// TIA Portal V20 export
DATA_BLOCK "POS3_0_Signal"   // DB34
{ S7_Optimized_Access := 'TRUE' }
// stored: MemoryReserve 100
   VAR
      Schrittkette { S7_SetPoint := 'True'} : "Schrittkettenaufruf";
      Station { S7_SetPoint := 'True'} : "Schrittkettensteuerung";
      "Richten nach Not Aus" : Bool := FALSE;
      Erster_Durchlauf : Bool := TRUE;
   END_VAR
   VAR RETAIN
      Taktzeit : Array[0..10] of Time;
   END_VAR
   VAR
      M_Zyklus_start : Bool := FALSE;
      M_Zyklus_ende : Bool := TRUE;
   END_VAR
   VAR RETAIN
      Sollzyklen : Int;
      Istzyklen : Int;
      Restzyklen : Int;
      "-1001T1 Oriental_Positionen" { S7_SetPoint := 'True'} : "Oriental_Variablen_Positionen";
      "-1001T1 Oriental_Steuerung" { S7_SetPoint := 'True'} : "Oriental_Variablen_Steuerung";
      "-1001T1 Oriental_Beschleunigung" : Real := 2.0;
      "-1001T1 Oriental_Speed" : Real := 2.0;
   END_VAR
   VAR
      "-1001T1 Oriental_E_P-Preset" : Bool;
   END_VAR
   VAR RETAIN
      "-1002T1 Oriental_Positionen" { S7_SetPoint := 'True'} : "Oriental_Variablen_Positionen";
      "-1002T1 Oriental_Steuerung" { S7_SetPoint := 'True'} : "Oriental_Variablen_Steuerung";
      "-1002T1_Oriental_Beschleunigung" : Real := 2.0;
      "-1002T1_Oriental_Speed" : Real := 2.0;
   END_VAR
   VAR
      "-1002T1 Oriental_E_P-Preset" : Bool;
   END_VAR
   VAR RETAIN
      "-1002T1 Oriental_Umdrehungszähler" : Real;
      "-1002T1 Oriental_Absolute_Position" : Real;
   END_VAR
   VAR
      "-1012B1 Kraftsensor" : Real;   // -1012B1 Kraftsensor
   END_VAR
   VAR RETAIN
      "-POS3_0_Regelventil_Ausgleichszylinder_Sollwert" : Int;   // +Feld-940RN1 Regelventil Ausgleichszylinder Sollwert in mbar
   END_VAR
   VAR
      "-POS3_0_Regelventil_Ausgleichszylinder_Istwert" : Int;   // +Feld-940RN1 Regelventil Ausgleichszylinder Istwert in mbar
   END_VAR
   VAR RETAIN
      "-POS3_0_Regelventil_Ausgleichszylinder_Maximale_Abweichung" : Int;   // +Feld-940RN1 Regelventil Ausgleichszylinder Istwert in mbar
   END_VAR
   VAR
      "-POS3_0_Regelventil_Ausgleichszylinder_Abweichung_OK" : Bool;   // +Feld-940RN1 Regelventil Ausgleichszylinder Istwert in mbar
   END_VAR
   VAR RETAIN
      "-POS3_0_Regelventil_Überlastzylinder_Sollwert" : Int;   // +Feld-940RN2 Regelventil Überlastzylinder Sollwert in mbar
   END_VAR
   VAR
      "-POS3_0_Regelventil_Überlastzylinder_Istwert" : Int;   // +Feld-940RN2 Regelventil Überlastzylinder Istwert in mbar
   END_VAR
   VAR RETAIN
      "-POS3_0_Regelventil_Überlastzylinder_Maximale_Abweichung" : Int;   // +Feld-940RN2 Regelventil Überlastzylinder Istwert in mbar
   END_VAR
   VAR
      "-POS3_0_Regelventil_Überlastzylinder_Abweichung_OK" : Bool;   // +Feld-940RN2 Regelventil Überlastzylinder Istwert in mbar
      "-POS3.0_Wegmessung_Ausgleichszylinder_Istwert_Rohwert" : Int;   // +POS=3.0-1011B1 Wegmessung Ausgleichszylinder Istwert Rohwert
   END_VAR
   VAR RETAIN
      "-POS3.0_Wegmessung_Ausgleichszylinder_Maximale_Abweichung" : Int;   // Wegmessung Ausgleichszylinder Toleranz in mm
      "-POS3.0_Wegmessung_Ausgleichszylinder_Position_GS_Abweichung_OK" : Bool;   // +POS=3.0-1011B1 Wegmessung Ausgleichszylinder Position GS Abweichung OK
      "-POS3.0_Wegmessung_Ausgleichszylinder_Position_AS1_Abweichung_OK" : Bool;   // +POS=3.0-1011B1 Wegmessung Ausgleichszylinder Position AS1 Abweichung OK
      Kommunikation_Weiterschaltbedingungen_AUS : Bool := 1;   // Kommunikation_Weiterschaltbedingungen_AUS
      Kommunikation_Weiterschaltbedingungen_DIGITAL : Bool;   // Kommunikation_Weiterschaltbedingungen_DIGITAL
      Kommunikation_Weiterschaltbedingungen_SP7 : Bool;   // Kommunikation_Weiterschaltbedingungen_SP7
   END_VAR
   VAR
      "-POS3.0_Wegmessung_Ausgleichszylinder_Sollwert_in_mm" : Real;   // +POS=3.0-1011B1 Wegmessung Ausgleichszylinder Sollwert in mm
      "-POS3.0_Wegmessung_Ausgleichszylinder_Istwert_in_mm" : Real;   // +POS=3.0-1011B1 Wegmessung Ausgleichszylinder Istwert in mm
   END_VAR
   VAR RETAIN
      "-POS3.0_Wegmessung_Ausgleichszylinder_Nullpunkt_Rohwert" : Int;   // +POS=3.0-1011B1 Wegmessung Ausgleichszylinder Nullpunkt Rohwert
   END_VAR
   VAR
      "-POS3.0_Wegmessung_Ausgleichszylinder_Taster_Nullen" : Bool;   // +POS=3.0-1011B1 Wegmessung Ausgleichszylinder Taster Nullen
   END_VAR
   VAR RETAIN
      "-POS3.0_Wegmessung_Ausgleichszylinder_Position_GS_aktiv" : Bool;   // +POS=3.0-1011B1 Wegmessung Ausgleichszylinder Position GS aktiv
      "-POS3.0_Wegmessung_Ausgleichszylinder_Position_AS1_aktiv" : Bool;   // +POS=3.0-1011B1 Wegmessung Ausgleichszylinder Position AS1 aktiv
      "Wartezeit Soll gesteckt" : Time;   // Wartezeit Soll gesteckt aus Verwaltung [s]
      "Wartezeit Ist gesteckt" : Real;   // Wartezeit Ist gesteckt für Anzeige [s]
   END_VAR
   VAR
      Status_gesteckt : Bool;   // Status Stecker ist gesteckt
      Drehachse_Kraft_überschritten : Bool;   // Drehachse Kraft überschritten
   END_VAR
BEGIN
   Schrittkette.OFF_SQ := FALSE;
   Schrittkette.INIT_SQ := FALSE;
   Schrittkette.ACK_EF := FALSE;
   Schrittkette.HALT_SQ := FALSE;
   Schrittkette.HALT_TM := FALSE;
   Schrittkette.ZERO_OP := FALSE;
   Schrittkette.EN_IL := FALSE;
   Schrittkette.EN_SV := FALSE;
   Schrittkette.S_PREV := FALSE;
   Schrittkette.S_NEXT := FALSE;
   Schrittkette.SW_AUTO := FALSE;
   Schrittkette.SW_TAP := FALSE;
   Schrittkette.SW_MAN := FALSE;
   Schrittkette.S_SEL := 0;
   Schrittkette.S_ON := FALSE;
   Schrittkette.S_OFF := FALSE;
   Schrittkette.T_PUSH := FALSE;
   Schrittkette.S_NO := 1;
   Schrittkette.S_MORE := FALSE;
   Schrittkette.S_ACTIVE := FALSE;
   Schrittkette.ERR_FLT := FALSE;
   Schrittkette.SQ_HALTED := FALSE;
   Schrittkette.TM_HALTED := FALSE;
   Schrittkette.OP_ZEROED := FALSE;
   Schrittkette.IL_ENABELD := FALSE;
   Schrittkette.SV_ENABELD := FALSE;
   Schrittkette.AUTO_ON := TRUE;
   Schrittkette.TAP_ON := FALSE;
   Schrittkette.MAN_ON := FALSE;
   Station.SK_Freigabe_Richten := FALSE;
   Station.SK_Richten_gestartet := FALSE;
   Station.SK_Richten_fertig := FALSE;
   Station.SK_Freigabe_Auto := FALSE;
   Station.SK_Aktiv := FALSE;
   Station.SK_Fertig := FALSE;
   Station.SK_Freigabe_Manuell_Auto := FALSE;
   Station.SK_Freigabe_Manuell_Richten := FALSE;
   Station.Reset_Freigaben := FALSE;
   Station.Station_1Ein_0Aus := FALSE;
   Station.SK_Richten_erforderlich := FALSE;
   Taktzeit[0..10] := T#0MS;
   "-1001T1 Oriental_Positionen".Start_POS_Position[0..15] := FALSE;
   "-1001T1 Oriental_Positionen".POS_OK_Position[0] := TRUE;
   "-1001T1 Oriental_Positionen".POS_OK_Position[1..15] := FALSE;
   "-1001T1 Oriental_Positionen".Operation_type[0..15] := 16#0001;
   "-1001T1 Oriental_Positionen".Soll_Position[0..15] := 0.0;
   "-1001T1 Oriental_Positionen".Geschwindigkeit[0] := 10.0;
   "-1001T1 Oriental_Positionen".Geschwindigkeit[1..4] := 2.0;
   "-1001T1 Oriental_Positionen".Geschwindigkeit[5..15] := 20.0;
   "-1001T1 Oriental_Positionen".Start_Rampe[0..4] := 2.0;
   "-1001T1 Oriental_Positionen".Start_Rampe[5..15] := 100.0;
   "-1001T1 Oriental_Positionen".Stopp_Rampe[0..4] := 2.0;
   "-1001T1 Oriental_Positionen".Stopp_Rampe[5..15] := 100.0;
   "-1001T1 Oriental_Positionen".Arbeitsstrom[0] := 10;
   "-1001T1 Oriental_Positionen".Arbeitsstrom[1..4] := 50;
   "-1001T1 Oriental_Positionen".Arbeitsstrom[5..15] := 1000;
   "-1001T1 Oriental_Positionen".Positioniertoleranz[0..15] := 0.01;
   "-1001T1 Oriental_Positionen".A_Softw_ES_min_mm := -0.5;
   "-1001T1 Oriental_Positionen".A_Softw_ES_max_mm := 10000.5;
   "-1001T1 Oriental_Positionen".A_Max_Speed_mm_s := 0;
   "-1001T1 Oriental_Positionen".A_Max_Beschleunigung_mm_s := 0;
   "-1001T1 Oriental_Positionen".A_Softw_ES_min_steps := 0.0;
   "-1001T1 Oriental_Positionen".A_Softw_ES_max_steps := 0.0;
   "-1001T1 Oriental_Steuerung".E_TRIG := FALSE;
   "-1001T1 Oriental_Steuerung"."E_TRIG-MODE" := FALSE;
   "-1001T1 Oriental_Steuerung"."E_ETO-CLR" := FALSE;
   "-1001T1 Oriental_Steuerung"."E_FW-JOG" := FALSE;
   "-1001T1 Oriental_Steuerung"."E_RV-JOG" := FALSE;
   "-1001T1 Oriental_Steuerung".E_START := FALSE;
   "-1001T1 Oriental_Steuerung".E_ZHOME := FALSE;
   "-1001T1 Oriental_Steuerung".E_STOP := FALSE;
   "-1001T1 Oriental_Steuerung".E_FREE := FALSE;
   "-1001T1 Oriental_Steuerung"."E_ALM-RST" := FALSE;
   "-1001T1 Oriental_Steuerung".E_DDO_Type := 16#0000;
   "-1001T1 Oriental_Steuerung".E_DDO_Pos := 0.0;
   "-1001T1 Oriental_Steuerung".E_DDO_Vel := 2.0;
   "-1001T1 Oriental_Steuerung".E_DDO_Acc := 100.0;
   "-1001T1 Oriental_Steuerung".E_DDO_Dec := 100.0;
   "-1001T1 Oriental_Steuerung".E_DDO_Crnt := 16#0064;
   "-1001T1 Oriental_Steuerung".E_DDO_Trans := 16#0000;
   "-1001T1 Oriental_Steuerung".A_TRIG_R := FALSE;
   "-1001T1 Oriental_Steuerung"."A_TRIG-MODE_R" := FALSE;
   "-1001T1 Oriental_Steuerung"."A_SET-ERR" := FALSE;
   "-1001T1 Oriental_Steuerung"."A_EXE-ERR" := FALSE;
   "-1001T1 Oriental_Steuerung"."A_DCMD-FULL" := FALSE;
   "-1001T1 Oriental_Steuerung".A_STOP_R := FALSE;
   "-1001T1 Oriental_Steuerung"."A_ETO-MON" := FALSE;
   "-1001T1 Oriental_Steuerung".A_TLC := FALSE;
   "-1001T1 Oriental_Steuerung"."A_SEQ-BSY" := FALSE;
   "-1001T1 Oriental_Steuerung".A_MOVE := FALSE;
   "-1001T1 Oriental_Steuerung"."A_IN-POS" := TRUE;
   "-1001T1 Oriental_Steuerung".A_START_R := FALSE;
   "-1001T1 Oriental_Steuerung"."A_HOME-END" := FALSE;
   "-1001T1 Oriental_Steuerung".A_READY := TRUE;
   "-1001T1 Oriental_Steuerung"."A_DCMD-RDY" := TRUE;
   "-1001T1 Oriental_Steuerung"."A_ALM-A" := FALSE;
   "-1001T1 Oriental_Steuerung".A_PresentAlarm := 16#0000;
   "-1001T1 Oriental_Steuerung".A_FBposition := 0.0;
   "-1001T1 Oriental_Steuerung".A_FBspeed := 0.0;
   "-1001T1 Oriental_Steuerung".A_CmdPosition := 0;
   "-1001T1 Oriental_Steuerung".A_TorqueMonitor := -17;
   "-1001T1 Oriental_Steuerung".A_CST_OpeCurrent := 16#01F4;
   "-1001T1 Oriental_Steuerung".A_Information := 16#0000_0000;
   "-1001T1 Oriental_Steuerung".A_StatusWord := 16#0000_0004;
   "-1001T1 Oriental_Steuerung".E_Trig_Manuell := FALSE;
   "-1001T1 Oriental_Steuerung".E_Schrittweite_pos := FALSE;
   "-1001T1 Oriental_Steuerung".E_Schrittweite_neg := FALSE;
   "-1001T1 Oriental_Steuerung".E_Schrittweite := 90.0;
   "-1002T1 Oriental_Positionen".Start_POS_Position[0..15] := FALSE;
   "-1002T1 Oriental_Positionen".POS_OK_Position[0] := TRUE;
   "-1002T1 Oriental_Positionen".POS_OK_Position[1..15] := FALSE;
   "-1002T1 Oriental_Positionen".Operation_type[0..15] := 16#0001;
   "-1002T1 Oriental_Positionen".Soll_Position[0..15] := 0.0;
   "-1002T1 Oriental_Positionen".Geschwindigkeit[0] := 10.0;
   "-1002T1 Oriental_Positionen".Geschwindigkeit[1..4] := 2.0;
   "-1002T1 Oriental_Positionen".Geschwindigkeit[5..15] := 20.0;
   "-1002T1 Oriental_Positionen".Start_Rampe[0..4] := 2.0;
   "-1002T1 Oriental_Positionen".Start_Rampe[5..15] := 100.0;
   "-1002T1 Oriental_Positionen".Stopp_Rampe[0..4] := 2.0;
   "-1002T1 Oriental_Positionen".Stopp_Rampe[5..15] := 100.0;
   "-1002T1 Oriental_Positionen".Arbeitsstrom[0] := 10;
   "-1002T1 Oriental_Positionen".Arbeitsstrom[1..4] := 50;
   "-1002T1 Oriental_Positionen".Arbeitsstrom[5..15] := 1000;
   "-1002T1 Oriental_Positionen".Positioniertoleranz[0..3] := 0.001;
   "-1002T1 Oriental_Positionen".Positioniertoleranz[4..15] := 0.01;
   "-1002T1 Oriental_Positionen".A_Softw_ES_min_mm := -0.5;
   "-1002T1 Oriental_Positionen".A_Softw_ES_max_mm := 10000.5;
   "-1002T1 Oriental_Positionen".A_Max_Speed_mm_s := 0;
   "-1002T1 Oriental_Positionen".A_Max_Beschleunigung_mm_s := 0;
   "-1002T1 Oriental_Positionen".A_Softw_ES_min_steps := 0.0;
   "-1002T1 Oriental_Positionen".A_Softw_ES_max_steps := 0.0;
   "-1002T1 Oriental_Steuerung".E_TRIG := FALSE;
   "-1002T1 Oriental_Steuerung"."E_TRIG-MODE" := FALSE;
   "-1002T1 Oriental_Steuerung"."E_ETO-CLR" := FALSE;
   "-1002T1 Oriental_Steuerung"."E_FW-JOG" := FALSE;
   "-1002T1 Oriental_Steuerung"."E_RV-JOG" := FALSE;
   "-1002T1 Oriental_Steuerung".E_START := FALSE;
   "-1002T1 Oriental_Steuerung".E_ZHOME := FALSE;
   "-1002T1 Oriental_Steuerung".E_STOP := FALSE;
   "-1002T1 Oriental_Steuerung".E_FREE := FALSE;
   "-1002T1 Oriental_Steuerung"."E_ALM-RST" := FALSE;
   "-1002T1 Oriental_Steuerung".E_DDO_Type := 16#0000;
   "-1002T1 Oriental_Steuerung".E_DDO_Pos := 0.0;
   "-1002T1 Oriental_Steuerung".E_DDO_Vel := 2.0;
   "-1002T1 Oriental_Steuerung".E_DDO_Acc := 100.0;
   "-1002T1 Oriental_Steuerung".E_DDO_Dec := 100.0;
   "-1002T1 Oriental_Steuerung".E_DDO_Crnt := 16#0064;
   "-1002T1 Oriental_Steuerung".E_DDO_Trans := 16#0000;
   "-1002T1 Oriental_Steuerung".A_TRIG_R := FALSE;
   "-1002T1 Oriental_Steuerung"."A_TRIG-MODE_R" := FALSE;
   "-1002T1 Oriental_Steuerung"."A_SET-ERR" := FALSE;
   "-1002T1 Oriental_Steuerung"."A_EXE-ERR" := FALSE;
   "-1002T1 Oriental_Steuerung"."A_DCMD-FULL" := FALSE;
   "-1002T1 Oriental_Steuerung".A_STOP_R := FALSE;
   "-1002T1 Oriental_Steuerung"."A_ETO-MON" := FALSE;
   "-1002T1 Oriental_Steuerung".A_TLC := FALSE;
   "-1002T1 Oriental_Steuerung"."A_SEQ-BSY" := FALSE;
   "-1002T1 Oriental_Steuerung".A_MOVE := FALSE;
   "-1002T1 Oriental_Steuerung"."A_IN-POS" := TRUE;
   "-1002T1 Oriental_Steuerung".A_START_R := FALSE;
   "-1002T1 Oriental_Steuerung"."A_HOME-END" := FALSE;
   "-1002T1 Oriental_Steuerung".A_READY := TRUE;
   "-1002T1 Oriental_Steuerung"."A_DCMD-RDY" := TRUE;
   "-1002T1 Oriental_Steuerung"."A_ALM-A" := FALSE;
   "-1002T1 Oriental_Steuerung".A_PresentAlarm := 16#0000;
   "-1002T1 Oriental_Steuerung".A_FBposition := 0.0;
   "-1002T1 Oriental_Steuerung".A_FBspeed := 0.0;
   "-1002T1 Oriental_Steuerung".A_CmdPosition := 0;
   "-1002T1 Oriental_Steuerung".A_TorqueMonitor := -17;
   "-1002T1 Oriental_Steuerung".A_CST_OpeCurrent := 16#01F4;
   "-1002T1 Oriental_Steuerung".A_Information := 16#0000_0000;
   "-1002T1 Oriental_Steuerung".A_StatusWord := 16#0000_0004;
   "-1002T1 Oriental_Steuerung".E_Trig_Manuell := FALSE;
   "-1002T1 Oriental_Steuerung".E_Schrittweite_pos := FALSE;
   "-1002T1 Oriental_Steuerung".E_Schrittweite_neg := FALSE;
   "-1002T1 Oriental_Steuerung".E_Schrittweite := 90.0;
END_DATA_BLOCK
